(* Sampler test double that counts its calls and can be told to drop spans on start and to
   try to sample them again on end. *)
FUNCTION_BLOCK FB_Sampler_ForInspection EXTENDS FB_Sampler
VAR_INPUT
	dropOnStart: BOOL;  // clear the sampled bit in onStart
	sampleOnEnd: BOOL;  // set the sampled bit in onEnd
END_VAR
VAR_OUTPUT
	startCount: UDINT;
	endCount: UDINT;
END_VAR

METHOD onStart
VAR_INPUT
	span: REFERENCE TO FB_Span;
END_VAR
THIS^.startCount := THIS^.startCount + 1;
SUPER^.onStart(span:=span);
IF THIS^.dropOnStart THEN
	span.setSampled(FALSE);
END_IF
END_METHOD

METHOD onEnd
VAR_INPUT
	span: REFERENCE TO FB_Span;
END_VAR
THIS^.endCount := THIS^.endCount + 1;
IF THIS^.sampleOnEnd THEN
	span.setSampled(TRUE);
END_IF
END_METHOD

END_FUNCTION_BLOCK

(* stored: Version 1.1.0.1
   POU FB_Sampler_ForInspection: Id {6b42640f-b420-4746-9a33-dcb83742479f}, SpecialFunc None
   Method onStart: Id {22ae475f-7bf7-4866-89e6-05e57fe578e7}
   Method onEnd: Id {b16b0db0-b370-4093-93f9-4ea352af9b79} *)
